Fanuc KAREL source: compact_preamble.KL

PROGRAM NC0064
%NOLOCKGROUP
ROUTINE R
VAR
S1:INTEGER;S2:INTEGER;S3:INTEGER;S4:INTEGER
BEGIN
S1=1
FOR S2=1 TO 2 DO
FOR S3=1 TO 2 DO
FOR S4=1 TO 2 DO
S1=(S1 + 1)
ENDFOR
ENDFOR
ENDFOR
END R
BEGIN
R
END NC0064
